(*
	Processor test double that exposes the batch processor's record queue for assertions.
	Unlike FB_LogRecordProcessor_ForRecordsInspection it does NOT override
	onEmit, so tests exercise the real batch grouping behavior.
*)
FUNCTION_BLOCK FB_LogRecordProcessor_ForBatchInspection EXTENDS FB_LogRecordProcessor_Batch

// explicitly run the batch processor body so tests exercise the flush logic
SUPER^();

PROPERTY records : REFERENCE TO FB_LogRecordQueue
GET
records REF= THIS^._records;
END_GET
END_PROPERTY

END_FUNCTION_BLOCK

(* stored: Version 1.1.0.1
   POU FB_LogRecordProcessor_ForBatchInspection: Id {77cf6308-3d1f-410d-950d-b1dca7c648b7}, SpecialFunc None
   Property records: Id {f123a485-0b0c-4d1a-a6b7-26aed6beabce}
   Get Get: Id {f907df37-cc42-4b7f-92c6-7c91c79a1e96} *)
